(* IEC 61131-3 sources: daoli-st-library/_quarantine/R78, 4 files *)

(* ---- FC_DL_PressureUnitConvert.st ---- *)
(*==============================================================================
 * 组件名称 : FC_DL_PressureUnitConvert ｜ 子库 : DL_MathData ｜ v1.0.0 ｜ 2026-11-23
 * 平台     : CODESYS 3.5 / TwinCAT 3 / InoProShop / Machine Expert（纯 IEC，无厂商库）
 * 功能简介 : 压力单位 kPa / Bar / Psi / MPa 两两互转。源/目标由枚举对单向
 *            选择，单向基准链（先归一到 kPa）使公式域固定为 4+4 条分支。
 * 契约     : 返回换算结果 [目标单位]；枚举非法（越界值）返回 0.0；
 *            除数为编译期非零常量，无除零风险；纯函数无状态。
 * 依赖     : 无 DL_ 内部依赖（本批自足实现）
 * 红线自检 : R1 零全局 R2 零%I/%Q R3 纯IEC R4 枚举越界拒收返 0 + 常量除数
 *            R5 全变量与枚举项双语同行注释 R6 N/A（无状态机） R7 N/A
 * 修订历史 : 2026-11-23 R78-B1 工程单位换算族模板派生首版
 *============================================================================*)
TYPE E_DL_PressureUnit :
(
    eKPa := 0,      // 千帕 [kPa] / Kilo-pascal
    eBar,           // 巴 [bar] / Bar
    ePsi,           // 磅每平方英寸 [psi] / Pound per square inch
    eMPa            // 兆帕 [MPa] / Mega-pascal
);
END_TYPE

FUNCTION FC_DL_PressureUnitConvert : REAL
VAR_INPUT
    fValue : REAL;              // 输入数值 [源单位] / Input value in source unit
    eSrc : E_DL_PressureUnit;   // 源单位选择 / Source unit selector
    eDst : E_DL_PressureUnit;   // 目标单位选择 / Destination unit selector
END_VAR
VAR
    fBase : REAL;               // 归一化中间值 [kPa] / Normalized intermediate in kPa
END_VAR
FC_DL_PressureUnitConvert := 0.0;   // 缺省返回 0 / Default return 0
CASE eSrc OF                        // 段 1：归一到基准 kPa / Normalize to base kPa
    E_DL_PressureUnit.eKPa: fBase := fValue;                    // 基准直通 / Base pass-through
    E_DL_PressureUnit.eBar: fBase := fValue * 100.0;            // 1 bar = 100 kPa
    E_DL_PressureUnit.ePsi: fBase := fValue * 6.894757;         // 1 psi = 6.894757 kPa
    E_DL_PressureUnit.eMPa: fBase := fValue * 1000.0;           // 1 MPa = 1000 kPa
    ELSE FC_DL_PressureUnitConvert := 0.0; RETURN;              // 源枚举非法返 0 / Invalid source returns 0
END_CASE
CASE eDst OF                        // 段 2：基准到目标 / Base to destination
    E_DL_PressureUnit.eKPa: FC_DL_PressureUnitConvert := fBase;             // 基准直通 / Base pass-through
    E_DL_PressureUnit.eBar: FC_DL_PressureUnitConvert := fBase / 100.0;     // kPa 到 bar
    E_DL_PressureUnit.ePsi: FC_DL_PressureUnitConvert := fBase / 6.894757;  // kPa 到 psi
    E_DL_PressureUnit.eMPa: FC_DL_PressureUnitConvert := fBase / 1000.0;    // kPa 到 MPa
    ELSE FC_DL_PressureUnitConvert := 0.0;                      // 目标枚举非法返 0 / Invalid destination returns 0
END_CASE
END_FUNCTION

(* ---- FC_DL_QuantizeStepReal.st ---- *)
(*==============================================================================
 * 组件名称 : FC_DL_QuantizeStepReal ｜ 子库 : DL_MathData ｜ v1.0.0 ｜ 2026-11-23
 * 平台     : CODESYS 3.5 / TwinCAT 3 / InoProShop / Machine Expert（纯 IEC，无厂商库）
 * 功能简介 : 实数量化到 fStep 步距网格：吸附到最近的格点（nStep 倍数）。
 *            先除到步距域，经标准就近舍入型转换 REAL_TO_DINT 取最近
 *            格点序号，再映射回步距域。
 * 契约     : 返回量化后的网格值；fStep <= 0 或输入 NaN/Inf 恒返回 0.0；
 *            商超出 DINT 安全域时按原值近直返；纯函数无状态。
 * 依赖     : 无 DL_ 内部依赖（本批自足实现）
 * 红线自检 : R1 零全局 R2 零%I/%Q R3 纯IEC（*_TO_* 显式转换）R4 非法步距/
 *            NaN/Inf 返 0 + 商域闸防转换溢出 R5 双语注释
 *            R6 N/A（无状态机） R7 N/A（无定时器实例）
 * 修订历史 : 2026-11-23 R78-B1 对齐取整族模板派生首版
 *============================================================================*)
FUNCTION FC_DL_QuantizeStepReal : REAL
VAR_INPUT
    fValue : REAL;          // 输入实数 / Input real value
    fStep : REAL;           // 量化步距，须 > 0 / Quantization step, must be > 0
END_VAR
VAR
    fQ : REAL;              // 步距域商 / Ratio in step domain
    nQ : DINT;              // 最近格点序号 / Nearest grid index
END_VAR
VAR CONSTANT
    DL_Q_SAFE_MAX : REAL := 2.0E9;      // DINT 安全商上限，防转换溢出 / Safe ratio cap guarding conversion overflow
END_VAR
IF (fStep <= 0.0) OR (fValue <> fValue) OR ((fValue - fValue) <> 0.0) THEN
    FC_DL_QuantizeStepReal := 0.0;      // 非法步距或 NaN/Inf 输入返 0 / Invalid step or NaN/Inf returns 0
    RETURN;
END_IF
fQ := fValue / fStep;                           // 商 / Ratio
IF (fQ <> fQ) OR ((fQ - fQ) <> 0.0) OR (fQ > DL_Q_SAFE_MAX) OR (fQ < -DL_Q_SAFE_MAX) THEN
    FC_DL_QuantizeStepReal := fQ * fStep;       // 商 NaN/Inf/超域按原值近直返 / NaN/Inf/out-of-domain ratio returns near-original
    RETURN;
END_IF
nQ := REAL_TO_DINT(fQ);                         // 最近邻取整（IEC 实转整为就近舍入）/ Round to nearest via typed conversion
FC_DL_QuantizeStepReal := DINT_TO_REAL(nQ) * fStep;     // 映射回步距域 / Map back to step domain
END_FUNCTION

(* ---- FC_DL_RoundToMultipleInt.st ---- *)
(*==============================================================================
 * 组件名称 : FC_DL_RoundToMultipleInt ｜ 子库 : DL_MathData ｜ v1.0.0 ｜ 2026-11-23
 * 平台     : CODESYS 3.5 / TwinCAT 3 / InoProShop / Machine Expert（纯 IEC，无厂商库）
 * 功能简介 : 整数四舍五入到 nMultiple 的最近倍数（半值远离零舍入，
 *            Round Half Away From Zero）。纯整数算术实现，先向零截断得
 *            基准倍数，再按"余量是否过半"进位 / 退位，无浮点精度损失。
 * 契约     : 返回四舍五入后的倍数值；nMultiple <= 0 恒返回 0；
 *            纯函数无状态、同输入同输出。
 * 依赖     : 无 DL_ 内部依赖（本批自足实现）
 * 红线自检 : R1 零全局 R2 零%I/%Q R3 纯IEC R4 非法倍数返 0 + 比较用 nHalf
 *            避免 nRem*2 溢出 R5 双语注释 R6 N/A（无状态机） R7 N/A
 * 修订历史 : 2026-11-23 R78-B1 对齐取整族模板派生首版
 *============================================================================*)
FUNCTION FC_DL_RoundToMultipleInt : DINT
VAR_INPUT
    nValue : DINT;          // 输入整数 / Input integer value
    nMultiple : DINT;       // 对齐倍数，须 > 0 / Alignment multiple, must be > 0
END_VAR
VAR
    nLo : DINT;             // 向零截断的基准倍数值 / Truncated-toward-zero base multiple
    nRem : DINT;            // 余量，符号随被除数，绝对值 < nMultiple / Remainder, |nRem| < nMultiple
    nHalf : DINT;           // 倍数半值（向下取整） / Floor half of the multiple
END_VAR
IF nMultiple <= 0 THEN
    FC_DL_RoundToMultipleInt := 0;      // 非法倍数返 0 / Invalid multiple returns 0
    RETURN;
END_IF
nLo := (nValue / nMultiple) * nMultiple;    // 整除截取得基准 / Base via integer division truncation
nRem := nValue - nLo;                       // 余量 / Remainder in (-nMultiple, nMultiple)
nHalf := nMultiple / 2;                     // 半值基准，免 nRem*2 溢出 / Half reference avoids nRem*2 overflow
IF nRem >= 0 THEN
    IF (nRem > nHalf) OR ((nRem = nHalf) AND ((nMultiple MOD 2) = 0)) THEN
        nLo := nLo + nMultiple;             // 正余量过半进位 / Round up at half
    END_IF
ELSIF (-nRem > nHalf) OR ((-nRem = nHalf) AND ((nMultiple MOD 2) = 0)) THEN
    nLo := nLo - nMultiple;                 // 负余量过半退位 / Round down at half
END_IF
FC_DL_RoundToMultipleInt := nLo;            // 输出四舍五入结果 / Output rounded result
END_FUNCTION

(* ---- FC_DL_SnapToStepLreal.st ---- *)
(*==============================================================================
 * 组件名称 : FC_DL_SnapToStepLreal ｜ 子库 : DL_MathData ｜ v1.0.0 ｜ 2026-11-23
 * 平台     : CODESYS 3.5 / TwinCAT 3 / InoProShop / Machine Expert（纯 IEC，无厂商库）
 * 功能简介 : LREAL 吸附到 fStep 步距网格的最近格点。双精度版量化件：
 *            先除到步距域，经标准就近舍入型转换 LREAL_TO_LINT 取最近
 *            格点序号（64 位序号域），再映射回步距域。
 * 契约     : 返回吸附后的网格值 [fStep 单位]；fStep <= 0 或输入 NaN 恒
 *            返回 0.0；商为 Inf 或超出 LINT 安全域时按原值近直返；
 *            纯函数无状态、同输入同输出。
 * 依赖     : 无 DL_ 内部依赖（本批自足实现）
 * 红线自检 : R1 零全局 R2 零%I/%Q R3 纯IEC（*_TO_* 显式转换）R4 非法步距/
 *            NaN 返 0 + 商域闸防转换溢出 R5 双语注释
 *            R6 N/A（无状态机） R7 N/A（无定时器实例）
 * 修订历史 : 2026-11-23 R78-B1 对齐取整族模板派生首版
 *============================================================================*)
FUNCTION FC_DL_SnapToStepLreal : LREAL
VAR_INPUT
    fValue : LREAL;         // 输入双精度实数 / Input LREAL value
    fStep : LREAL;          // 量化步距，须 > 0 / Quantization step, must be > 0
END_VAR
VAR
    fQ : LREAL;             // 步距域商 / Ratio in step domain
    nQ : LINT;              // 最近格点序号（64 位域） / Nearest grid index (64-bit domain)
END_VAR
VAR CONSTANT
    DL_Q_SAFE_MAX : LREAL := 9.0E18;    // LINT 安全商上限，防转换溢出 / Safe ratio cap guarding conversion overflow
END_VAR
IF (fStep <= 0.0) OR (fValue <> fValue) OR ((fValue - fValue) <> 0.0) THEN
    FC_DL_SnapToStepLreal := 0.0;       // 非法步距或 NaN 输入返 0 / Invalid step or NaN returns 0
    RETURN;
END_IF
fQ := fValue / fStep;                           // 商 / Ratio
IF (fQ <> fQ) OR ((fQ - fQ) <> 0.0) OR (fQ > DL_Q_SAFE_MAX) OR (fQ < -DL_Q_SAFE_MAX) THEN
    FC_DL_SnapToStepLreal := fQ * fStep;        // 商 NaN/Inf/超域按原值近直返 / NaN/Inf/out-of-domain ratio returns near-original
    RETURN;
END_IF
nQ := LREAL_TO_LINT(fQ);                        // 最近邻取整（IEC 实转整为就近舍入）/ Round to nearest via typed conversion
FC_DL_SnapToStepLreal := LINT_TO_LREAL(nQ) * fStep;     // 映射回步距域 / Map back to step domain
END_FUNCTION
